Staubli VAL3: click_End.pgx

program click_End()
  local bool l_bResult
begin
   //循环停止机器人
  l_bResult=userPageConfirm("确认循环停止机器人？")
  if l_bResult
    rs:nCycleCmd=5
    delay(0.2)
    rs:nCycleCmd=0
  endIf
end
